FUNCTION FC 1 : VOID
BEGIN
NETWORK
      L 'AB
END_FUNCTION
